// TIA Portal V18 export
VAR_GLOBAL   // PLC tag table "LEITOR_VIVERK"
   Readcomplete AT %I2000.1 : Bool;
   ResultData0 AT %IB2284 : Byte;
   ResultData1 AT %IB2285 : Byte;
   ResultData2 AT %IB2286 : Byte;
   ResultData3 AT %IB2287 : Byte;
   ResultData4 AT %IB2288 : Byte;
   ResultData5 AT %IB2289 : Byte;
   ResultData6 AT %IB2290 : Byte;
   ResultData7 AT %IB2291 : Byte;
   ResultData8 AT %IB2292 : Byte;
   ResultData9 AT %IB2293 : Byte;
   ResultData10 AT %IB2294 : Byte;
   ResultData11 AT %IB2295 : Byte;
   ResultData12 AT %IB2296 : Byte;
   Tag_5 AT %IB2000 : Byte;
   Tag_6 AT %IB2001 : Byte;
   Tag_7 AT %IB2002 : Byte;
   Tag_8 AT %IB2003 : Byte;
   Tag_9 AT %IB2004 : Byte;
   Tag_10 AT %IB2005 : Byte;
   Tag_11 AT %IB2006 : Byte;
   Tag_12 AT %IB2007 : Byte;
   Tag_13 AT %IB2008 : Byte;
   Tag_14 AT %IB2009 : Byte;
   Tag_15 AT %IB2010 : Byte;
   Tag_16 AT %IB2011 : Byte;
   Tag_17 AT %IB2012 : Byte;
   Tag_18 AT %IB2013 : Byte;
END_VAR
